RoboDK station: pick and place.rdk

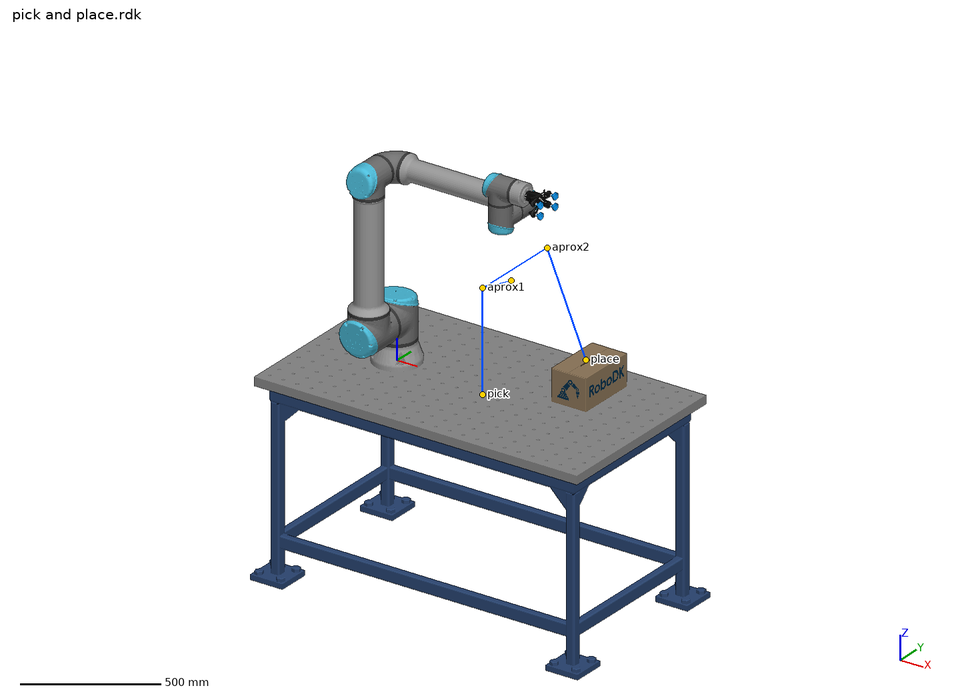
[picture v0: the station drawn from its stored meshes, robots at their saved joint values, targets as dots, program paths as lines]
Station Nueva Estación (1) (saved by RoboDK 6.2.0). Poses are relative to the parent item; angles as X-Y-Z fixed-axis rotations.
  - frame UR10e Base at (0, 0, 0) mm
    - robot UR10e: 6 axes, payload 10 kg, reach 1300 mm, repeatability 0.05 mm, weight 28.9 kg
        modified DH rows (alpha deg, a mm, theta deg, d mm): 0, 0, 0, 180.7; 90, 0, 180, 0; 0, 612.6, 0, 0; 0, 571.335, 0, 174.15; -90, 0, 0, 119.85; 90, 0, 180, 116.55
        joint limits [-360, -360, -360, -360, -360, -360] to [360, 360, 360, 360, 360, 360]; home [0, -90, -90, 0, 90, 0]; saved at [0, -90, -90, 0, 90, 0]
      - tool RobotiQ EPick Vacuum Gripper (4 Cups), TCP at (0, 15, 90) mm, size 119.5 x 73.5 x 92.5 mm
    - target pick (Cartesian target) at (560, -270, 130) mm, rotated rx 180 ry 0 rz 90 deg; joints [-9.716, -100.097, -131.425, -38.477, 89.999, -189.716] of UR10e
    - target aprox1 (Cartesian target) at (560, -270, 550) mm, rotated rx 180 ry 0 rz 90 deg; joints [-9.716, -79.865, -102.863, -87.27, 89.999, -189.716] of UR10e
    - target aprox2 (Cartesian target) at (560, 130, 550) mm, rotated rx 180 ry 0 rz 90 deg; joints [31.526, -75.012, -106.584, -88.404, 89.998, -148.474] of UR10e
    - target place (Cartesian target) at (700, 170, 130) mm, rotated rx 180 ry 0 rz 90 deg; joints [28.223, -107.635, -120.874, -41.491, 89.998, -151.777] of UR10e
    - target home (Cartesian target) at (682.46, -266.51, 612.24) mm, rotated rx 180 ry 0 rz -90 deg; joints [-7.424, -93.32, -84.019, -92.661, 90, -7.424] of UR10e
  - Python program Prog1 (listed below)
  - object Table 1400x800x800mm at (0, 0, 0) mm, size 1420 x 820 x 800 mm, geometry from Table-1400x800x800mm.sld
  - program Prog2 (12 instructions, listed below)
  - object Box 20x12in (Closed) at (640, 40, 0) mm, size 151.4 x 254.3 x 133.7 mm, geometry from Box-20x12in-Closed.sld
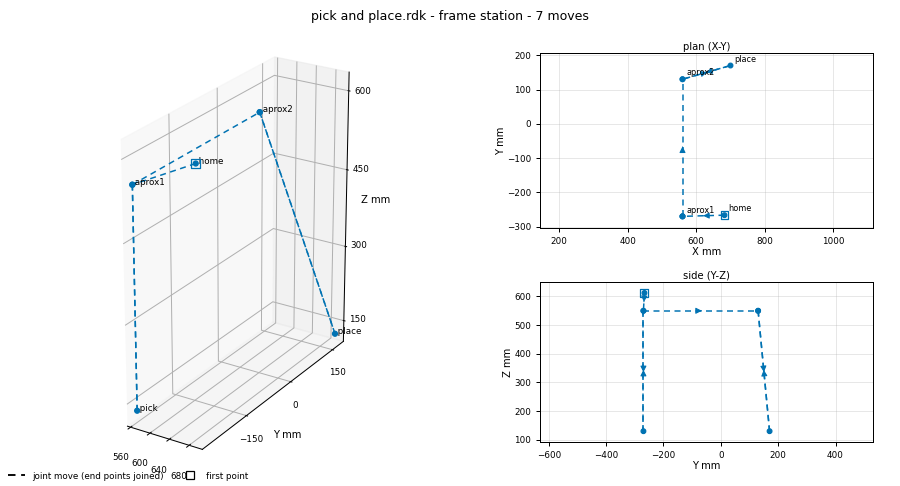
[picture p0: tool path of pick and place.rdk in frame station, 7 of 7 moves have a stored position in this frame; points joined in program order, loops and branches not executed]

--- Python program Prog1 ---
from robodk.robolink import *

RDK = Robolink()
robot = RDK.Item('UR10', ITEM_TYPE_ROBOT)

robot.MoveJ([0, -90, -90, 0, 90, 0])     # posición inicial
robot.MoveJ([45, -90, -90, 0, 90, 0])    # gira la base 45°
robot.MoveJ([-45, -90, -90, 0, 90, 0])   # gira la base al otro lado
robot.MoveJ([0, -90, -90, 0, 90, 0])     # vuelve al inicio

--- program Prog2 (robot UR10e) ---
  Est. Ref.: UR10e Base
  Est. herr: RobotiQ EPick Vacuum Gripper (4 Cups)
  Mover Box 20x12in (Closed)
  MoveJ (home)
  MoveJ (aprox1)
  MoveJ (pick)
  Adjuntar a RobotiQ EPick Vacuum Gripper (4 Cups)
  MoveJ (aprox1)
  MoveJ (aprox2)
  MoveJ (place)
  Separar de RobotiQ EPick Vacuum Gripper (4 Cups)
  MoveJ (aprox2)
